Fanuc KAREL source: ko00059.KL

-- PROVISIONAL review KL for V1013-1; original PC SHA256 edfb7f41e2ea626a4b8e40306485abeb64013847f90dd67a9762db5bc031fbbb
-- Incomplete behavior may be omitted. Consult companion uncertainty JSON. Do not deploy.
PROGRAM KO00059
%NOLOCKGROUP
BEGIN
  -- UNRESOLVED_PC offsets 5-12; opcodes 9D,23
  -- UNRESOLVED_PC offsets 17-69; opcodes 27,27,49,7E,AD,27,49,7E,AD,22,31,7E,4A
  -- UNRESOLVED_PC offsets 74-78; opcodes 7F
END KO00059
